(* Tests that the file log exporter writes processed batches to disk. *)
FUNCTION_BLOCK FB_TestFileExporter EXTENDS FB_TestSuite
VAR
	_resource:		FB_Resource(schemaUrl:='');
	_exporter: 		FB_LogRecordExporter_File(filepath:='C:\Users\samue\Desktop\programming projects\TcOtlp\logs.jsonl');
	_processor:		FB_LogRecordProcessor_ForRecordsInspection(
		maxQueueSize:=0,
		scheduledDelayMillis:=1000,
		maxExportBatchSize:=512,
		exporter:=0
	);
	_provider:		FB_LoggerProvider(resource:=_resource);
	_scope1:			FB_InstrumentationScope(name:='scope1', version:='0.0.1', schemaUrl:='');
	_logger1:		FB_Logger(scope:=_scope1, provider:=_provider);
	_scope2:			FB_InstrumentationScope(name:='scope2', version:='0.0.1', schemaUrl:='');
	_logger2:		FB_Logger(scope:=_scope2, provider:=_provider);
END_VAR

THIS^.testExportBatchedLogRecords(cleanup:=FALSE);

(*
	Records emitted through two loggers reach the file as one batch, and a batch handed over in the
	scan the previous one finished still starts, so back-to-back flushes never stall the file exporter.
*)
METHOD testExportBatchedLogRecords : REFERENCE TO FB_Test

VAR_INPUT
	cleanup: BOOL := TRUE;  // FALSE keeps logs.jsonl on disk for manual inspection
END_VAR

VAR CONSTANT
	_filepath: STRING := 'C:\Users\samue\Desktop\programming projects\TcOtlp\logs.jsonl';
	MAX_CYCLES: UDINT := 1000;
END_VAR

VAR_INST
	_cycles: 		UDINT;
	_state:			USINT;
	_redelivered:	BOOL;  // a second batch was exported in the scan the first finished
	_fileFinder: 	FB_EnumFindFileEntry;
	_fileDeleter:	FB_FileDelete;
END_VAR

VAR
	_num: UINT;
	_fileSize: ULINT;
	_exportSucceeded: BOOL;
	_exportCallSucceeded: BOOL;
	_firstEmitSucceeded: BOOL;
	_secondEmitSucceeded: BOOL;
	_thirdEmitSucceeded: BOOL;
	_loggerFailureResult: E_LoggerFailureReason;
	_exporterFailureReason: E_LogRecordExporterFailureReason;
	_timestamp: ULINT := ULINT#1581452773000000789;
	_traceId: ARRAY[0..ValueFactory.nTraceIdBytes-1] OF BYTE := [0, 1, 2, 3, 4, 5, 6, 7, 8, 9, 10, 11, 12, 13, 14, 15];
	_spanId: ARRAY[0..ValueFactory.nSpanIdBytes-1] OF BYTE := [16, 17, 18, 19, 20, 21, 22, 23];
END_VAR
TcUnit.TEST('testExportBatchedLogRecords');
	CASE _state OF
		0: // emit three records through two loggers; the processor captures them without exporting
			_cycles := 0;
			_redelivered := FALSE;
			_processor.free();
			_logger1.free();
			// _resource persists across test re-runs; only add the attribute once
			IF _resource.attributes.count = 0 THEN
				_resource.attributes.setStringAttribute('host.id', 'PLC1');
			END_IF
			_num := 1;
			_firstEmitSucceeded := _logger1
				.startLogRecord(severityNumber:=E_SeverityNumber.DEBUG)
				.setTimestamp(_timestamp)
				.setBody('First batched log record')
				.setEventName('BatchRecord1')
				._setTraceId(ADR(_traceId), SIZEOF(_traceId))
				._setSpanId(ADR(_spanId), SIZEOF(_spanId))
				.setStringAttribute('batch.position', 'first')
				.setNumberAttribute('batch.positionNum', _num)
				.emit(failureResult=>_loggerFailureResult);
			_num := 2;
			_secondEmitSucceeded := _logger2
				.startLogRecord(severityNumber:=E_SeverityNumber.INFO)
				.setTimestamp(_timestamp)
				.setBody('Second batched log record')
				.setEventName('BatchRecord2')
				.setStringAttribute('batch.position', 'second')
				.setNumberAttribute('batch.positionNum', _num)
				.emit(failureResult=>_loggerFailureResult);
			_num := 3;
			_thirdEmitSucceeded := _logger1
				.startLogRecord(severityNumber:=E_SeverityNumber.WARN)
				.setTimestamp(_timestamp)
				.setBody('Third batched log record')
				.setEventName('BatchRecord3')
				.setStringAttribute('batch.position', 'third')
				.setNumberAttribute('batch.positionNum', _num)
				.emit(failureResult=>_loggerFailureResult);
			_provider
				.stageProcessor(_processor)
				.tick();
			THIS^.AssertTrue(_firstEmitSucceeded, 'Expected the first emit to succeed');
			THIS^.AssertTrue(_secondEmitSucceeded, 'Expected the second emit to succeed');
			THIS^.AssertTrue(_thirdEmitSucceeded, 'Expected the third emit to succeed');
			THIS^.AssertTrue(_logger1.pLogRecord = 0, 'Expected emit to release the logger-owned record');
			IF _firstEmitSucceeded
				AND _secondEmitSucceeded
				AND _thirdEmitSucceeded THEN
				THIS^.AssertEquals_UDINT(3, _processor.records.count, 'Expected the processor to capture all three log records');
				_state := 10;
				RETURN;
			ELSE
				_state := 30;
				RETURN;
			END_IF
			
		10: // hand the captured records to the file exporter and tick it until the write is done
			IF _processor.records.count > 0 THEN
				_exportSucceeded := _processor.exportRecords(
					exporter:=_exporter,
					failureReason=>_exporterFailureReason
				);
				IF NOT _exportSucceeded OR_ELSE _processor.records.count > 0 THEN
					THIS^.AssertTrue(FALSE, 'Expected the exporter to take ownership of the processor buffer');
					_state := 30;
					RETURN;
				END_IF
			END_IF
			_exportCallSucceeded := _exporter.tick(failureReason=>_exporterFailureReason);
			_cycles := _cycles + 1;
			IF NOT _exportCallSucceeded THEN
				THIS^.AssertTrue(
					_exporterFailureReason <> E_LogRecordExporterFailureReason.NA,
					'Expected an exporter failure reason when tick returns FALSE'
				);
				THIS^.AssertTrue(FALSE, 'Expected the file export to succeed');
				_state := 30;
				RETURN;
			ELSIF _cycles > MAX_CYCLES THEN
				THIS^.AssertTrue(FALSE, 'Expected the file export to finish within MAX_CYCLES');
				_state := 30;
				RETURN;
			ELSIF _exporter.currentState = E_FileExporterState.done AND NOT _redelivered THEN
				// hand over the next batch in the same scan; the exporter must still start it
				_redelivered := TRUE;
				_logger2
					.startLogRecord(severityNumber:=E_SeverityNumber.INFO)
					.setTimestamp(_timestamp)
					.setBody('Batch exported the scan the previous one finished')
					.emit(failureResult=>_loggerFailureResult);
				_provider
					.stageProcessor(_processor)
					.tick();
				_exportSucceeded := _processor.exportRecords(
					exporter:=_exporter,
					failureReason=>_exporterFailureReason
				);
				THIS^.AssertTrue(_exportSucceeded, 'Expected the finished exporter to accept the next batch');
				RETURN;
			ELSIF _exporter.currentState = E_FileExporterState.done THEN
				THIS^.AssertFalse(_exporter.isBusy(), 'Expected the exporter to release its completed records');
				THIS^.AssertTrue(
					_exporterFailureReason = E_LogRecordExporterFailureReason.NA,
					'Expected no failure reason when file export succeeds'
				);
				_state := 20;
				RETURN;
			ELSE
				RETURN;
			END_IF
			
		20: // verify the exported batch made the file non-empty
			_fileFinder(
				sPathName:=_filepath,
				bExecute:=TRUE,
			);
			IF NOT _fileFinder.bBusy THEN
				_fileSize := ULARGE_TO_ULINT(_fileFinder.stFindFile.fileSize);
				THIS^.AssertTrue(_fileSize > 0, 'Expected a non-empty file');
				_state := 30;
			END_IF
			RETURN;
		
		30: // cleanup the file
			IF cleanup THEN
				_fileDeleter(
					sPathName:=_filepath,
					bExecute:=TRUE,
				);
				IF _fileDeleter.bBusy THEN
					RETURN;
				END_IF
			END_IF

			// clean up the record owned by the processor
			_processor.free();
			_logger1.free();
			THIS^.AssertTrue(_processor.records.count = 0, 'Expected the processor to be empty after cleanup');

			_state := 0;
			TcUnit.TEST_FINISHED();
	END_CASE
END_METHOD

END_FUNCTION_BLOCK

(* stored: Version 1.1.0.1
   POU FB_TestFileExporter: Id {652c2ccf-e368-4316-b865-a55144794447}, SpecialFunc None
   Method testExportBatchedLogRecords: Id {62c42b19-8451-4cb9-878c-1813787327e9} *)
